(*
SPDX-FileCopyrightText: © 2026 Oleksandr Tiutyk <trofimich@gmail.com>
SPDX-License-Identifier: MIT
License: https://opensource.org/license/mit
*)

(*!
<summary>Names the two runs and intervening cancellation in the file-manager reuse test.</summary>
<description>
Steps belong to one test scenario; values are not a serialized protocol. The first member is the initial
preparation step. Test completion and failure cleanup are tracked separately.
</description>
*)
{attribute 'qualified_only'}
{attribute 'strict'}
{attribute 'to_string'}
TYPE FILE_MANAGER_REUSE_TEST_STEP :
(
	START_FIRST_WRITE,
	CANCEL_AFTER_WRITE,
	RESET_AND_START_SECOND_FILE,
	CHECK_SECOND_FILE
);
END_TYPE

(* stored: Version 1.1.0.1
   DUT FILE_MANAGER_REUSE_TEST_STEP: Id {aeb02eda-eb82-4112-a140-d9def4d96e61} *)
